(* IEC 61131-3 sources: rusty/tests/lit/cfc/blocks/function_feedback, 2 files *)

(* ---- main.st ---- *)
FUNCTION main : DINT
    function_feedback.seed := 5;
    function_feedback();
    function_feedback();
    // return feeds its own in1: cycle 1 => 0 + 5, cycle 2 => 5 + 5
    // CHECK: acc = 10
    printf('acc = %d$N', function_feedback.acc);
END_FUNCTION

(* ---- myAdd.st ---- *)
FUNCTION myAdd : INT
    VAR_INPUT
        in1, in2: DINT;
    END_VAR

    VAR_OUTPUT
        myAddDoubled: DINT;
    END_VAR

    myAdd := in1 + in2;
    myAddDoubled := (in1 + in2) * 2;
END_FUNCTION
